SUBAPPLICATION Uebung_263_AX (* Kein Blockieren: alle 10ms neuer PWM-Wert (0/4096) auf Q1 mit RAMP 500ms, Lebenszeichen Q2 blinkt 5 Hz gleichmaessig *)
  (* Standard: 61499-2; Description: Copyright (c) 2026 Meisterschulen am Ostbahnhof This program and the accompanying materials are made available under the terms of the Eclipse Public License 2.0 which is available at https://www.eclipse.org/legal/epl-2.0/ SPDX-License-Identifier: EPL-2.0 *)
  (* Version 1.0, 2026-11-06, Franz Höpfinger, Meisterschulen am Ostbahnhof, initial API and implementation and/or initial documentation *)
  PACKAGE Uebungen;
  IMPORT logiBUS::io::DQ::logiBUS_DO::Output_Q1;
  IMPORT logiBUS::io::DQ::logiBUS_DO::Output_Q2;
  (* Documentation:
  Kein Blockieren beim PWM-Wertwechsel
   Alle 10 ms bekommt Q1 einen neuen Wert (0 / 4096) bei RAMP = T#500ms. Jede Rampe wird nach 10 ms abgebrochen, die neue startet sofort am Ist-Wert.
   Erwartung:
    - Q2 blinkt gleichmäßig mit 5 Hz, Life_Count zählt gleichmäßig. Das ist der eigentliche Test.
   - Q1 bewegt sich kaum: Er pendelt nur wenige Prozent um den Startwert. Das ist erwartet.
   - RAMPO_Count_Q1 bleibt (fast) bei 0, weil abgebrochene Rampen kein RAMPO melden.
    Stockt Q2 oder Life_Count, blockiert der Wertwechsel den Event-Thread (alte Firmware oder altes ELF).
  *)
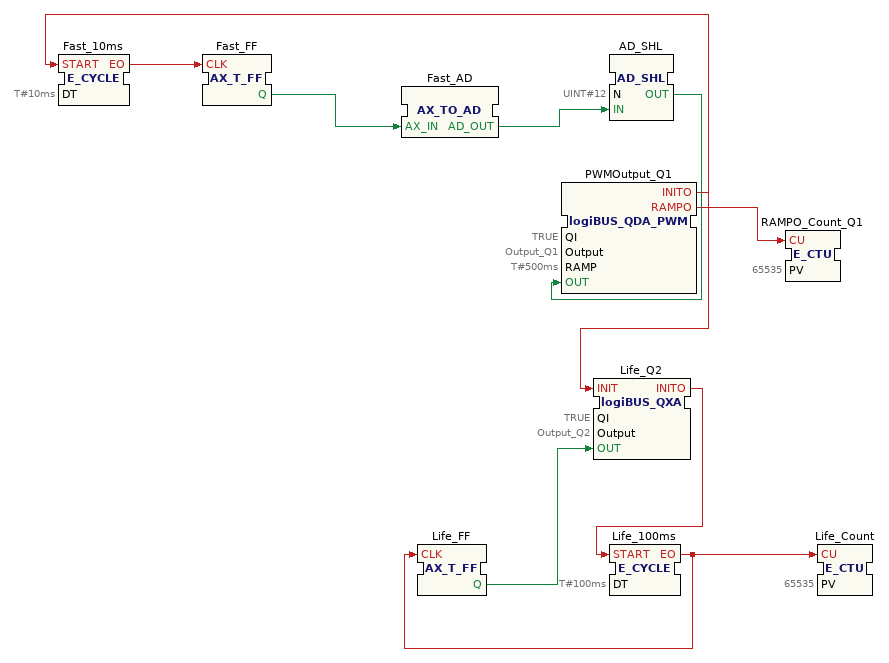
  FBS
    PWMOutput_Q1 : logiBUS::io::DQ::logiBUS_QDA_PWM(QI := TRUE, Output := Output_Q1, RAMP := T#500ms);
    Fast_10ms : iec61499::events::E_CYCLE(DT := T#10ms);
    Fast_FF : adapter::events::unidirectional::AX_T_FF;
    Fast_AD : adapter::conversion::unidirectional::AX_TO_AD;
    AD_SHL : adapter::iec61131::bitwise::AD_SHL(N := UINT#12);
    RAMPO_Count_Q1 : iec61499::events::E_CTU(PV := 65535);
    Life_100ms : iec61499::events::E_CYCLE(DT := T#100ms);
    Life_FF : adapter::events::unidirectional::AX_T_FF;
    Life_Q2 : logiBUS::io::DQ::logiBUS_QXA(QI := TRUE, Output := Output_Q2);
    Life_Count : iec61499::events::E_CTU(PV := 65535);
  END_FBS
  EVENT_CONNECTIONS
    PWMOutput_Q1.INITO TO Fast_10ms.START;
    Fast_10ms.EO TO Fast_FF.CLK;
    PWMOutput_Q1.RAMPO TO RAMPO_Count_Q1.CU;
    PWMOutput_Q1.INITO TO Life_Q2.INIT;
    Life_Q2.INITO TO Life_100ms.START;
    Life_100ms.EO TO Life_FF.CLK;
    Life_100ms.EO TO Life_Count.CU;
  END_CONNECTIONS
  ADAPTER_CONNECTIONS
    Fast_FF.Q TO Fast_AD.AX_IN;
    Life_FF.Q TO Life_Q2.OUT;
    Fast_AD.AD_OUT TO AD_SHL.IN;
    AD_SHL.OUT TO PWMOutput_Q1.OUT;
  END_CONNECTIONS
END_SUBAPPLICATION
